Fanuc KAREL source: ka00105.KL

PROGRAM KA00105
%STACKSIZE=65535
%PRIORITY=65535
%NOLOCKGROUP
VAR
SRC : VECTOR
DST : VECTOR
BEGIN
SRC.X=1.0
DST=SRC
END KA00105
